RESOURCE RES0 : EMB_RES_ECO
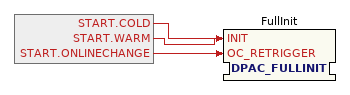
  FBS
    FullInit : DPAC_FULLINIT;
  END_FBS
  EVENT_CONNECTIONS
    START.COLD TO FullInit.INIT;
    START.WARM TO FullInit.INIT;
    START.ONLINECHANGE TO FullInit.OC_RETRIGGER;
  END_CONNECTIONS
END_RESOURCE
